Fanuc KAREL source: KT00738.KL

PROGRAM KT00738
%NOLOCKGROUP
VAR
  ARG: ARRAY[4] OF BYTE
  OUT: BOOLEAN
BEGIN
  OUT = UNINIT(ARG)
END KT00738
